RoboDK station: Bench V1 cell v4.rdk

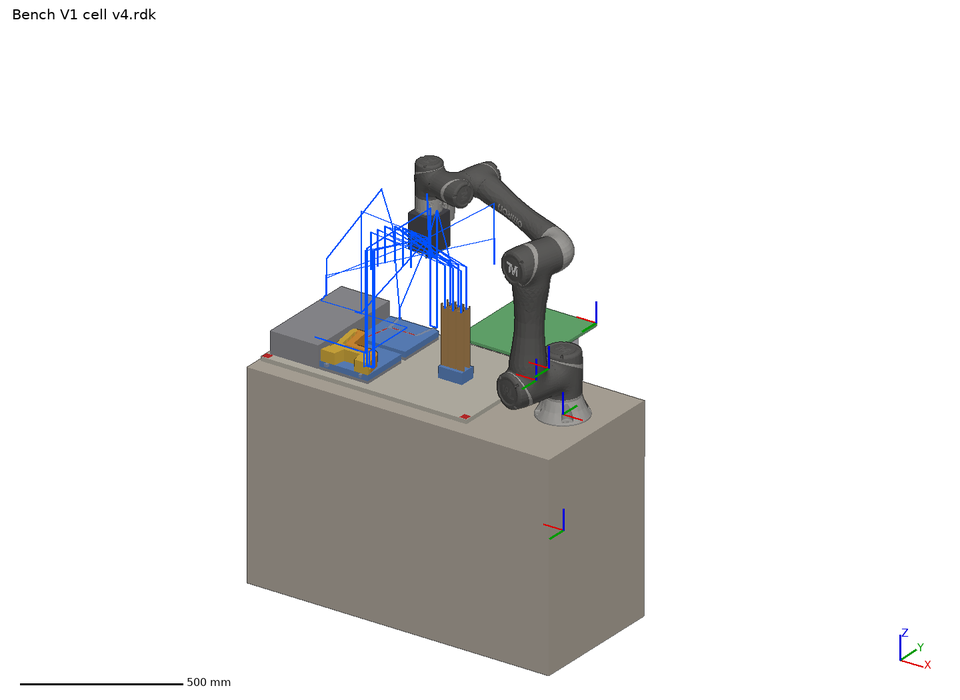
[picture v0: the station drawn from its stored meshes, robots at their saved joint values, targets as dots, program paths as lines]
Station Bench V1 cell v4 (saved by RoboDK 6.1.1). Poses are relative to the parent item; angles as X-Y-Z fixed-axis rotations.
Station parameters (name, value as stored): IO_0, 0
  - frame Cell at (0, 0, 0) mm
    - frame Work plate at (-206.44, 152.99, -4.46) mm, rotated rx -0.03 ry -0.07 rz -179.98 deg
      - frame Ground base at (0, -67, 15) mm
        - object Table at (0, 0, 0) mm, size 1130 x 510 x 735 mm
        - object Ground base plate at (0, 0, 0) mm, size 770 x 440 x 15 mm, geometry from ground_base_split.stl
        - object Vision square 1 at (3, 3, 0) mm, size 25 x 25 x 0.5 mm, geometry from vision_square.stl
        - object Vision square 2 at (742, 3, 0) mm, size 25 x 25 x 0.5 mm, geometry from vision_square.stl
        - object Vision square 3 at (3, 412, 0) mm, size 25 x 25 x 0.5 mm, geometry from vision_square.stl
        - object Vision square 4 at (742, 412, 0) mm, size 25 x 25 x 0.5 mm, geometry from vision_square.stl
        - object Base A riser at (480, 120, 10) mm, size 180 x 180 x 10 mm
        - object Base A at (480, 120, 10) mm, size 180 x 180 x 20 mm, geometry from base_a.stl
        - object Base B riser at (480, 320, 10) mm, size 180 x 180 x 10 mm
        - object Base B at (480, 320, 10) mm, size 180 x 180 x 20 mm, geometry from base_b.stl
        - object Plank jig at (150, 190, 0) mm, size 90 x 60 x 40 mm, geometry from plank_jig.stl
        - object Parking pad at (665, 220, 80) mm, size 180 x 380 x 80 mm, geometry from parking_pad.stl
        - frame AMR at (60, -340, 0) mm
          - object AMR plate at (0, 0, 0) mm, size 300 x 320 x 10 mm
          - object AMR top module at (0, 0, 0) mm, size 220 x 240 x 372 mm
          - frame Omron LD-250 Base at (150, -40, -765) mm
            - robot AMR LD-250: 4 axes
                joint limits [-10000, -10000, -10, -3600] to [10000, 10000, 10, 3600]; home [0, 0, 0, 0]; saved at [0, 0, 0, 0]
        - target Home (Cartesian target) at (295, 220, 380) mm, rotated rx 180 ry 0 rz 0 deg; joints [-14.089, 2.917, -80.099, -12.747, -90.01, 75.887] of Omron TM5-900
        - target guide B-A pick out low (Cartesian target) at (383, 390, 50) mm, rotated rx 0 ry 90 rz 0 deg; joints [8.389, -22.724, -132.74, -24.469, 98.365, 89.963] of Omron TM5-900
        - target guide B-A pick out (Cartesian target) at (383, 390, 450) mm, rotated rx 0 ry 90 rz 0 deg; joints [8.433, 10.061, -100.143, -89.851, 98.409, 89.963] of Omron TM5-900
        - target guide B-A via (Cartesian target) at (295, 220, 450) mm, rotated rx 0 ry 90 rz 0 deg; joints [-32.59, 30.389, -113.158, -97.152, 57.386, 90.016] of Omron TM5-900
        - target guide B-A centre (Cartesian target) at (295, 220, 450) mm, rotated rx 180 ry 0 rz 0 deg; joints [-14.088, -0.071, -66.923, -22.935, -90.01, 75.888] of Omron TM5-900
        - target guide B-A wrist ready (Cartesian target) at (295, 220, 450) mm, rotated rx -104.58 ry -32.51 rz -35.37 deg; joints [-50.735, 20.512, -106.829, -34.479, -14.275, 24.972] of Omron TM5-900
        - target guide B-A wrist swapped (joint target) at (338.92, 166.34, 566.06) mm, rotated rx -75.5 ry -32.53 rz -66.11 deg; joints [-50.735, 20.512, -106.829, -34.479, 14.275, 24.972] of Omron TM5-900
        - target guide B-A via (Cartesian target) at (295, 220, 450) mm, rotated rx 0 ry 90 rz 0 deg; joints [-32.59, 30.389, -113.158, -97.152, 57.386, 90.016] of Omron TM5-900
        - target guide B-A pick (Cartesian target) at (408, 390, 50) mm, rotated rx 0 ry 90 rz 0 deg; joints [7.812, -24.505, -129.214, -26.214, 97.788, 89.964] of Omron TM5-900
        - target guide B-A lift (Cartesian target) at (408, 390, 70) mm, rotated rx 0 ry 90 rz 0 deg; joints [7.814, -21.463, -128.95, -29.52, 97.79, 89.964] of Omron TM5-900
        - target guide B-A up (Cartesian target) at (408, 390, 450) mm, rotated rx 0 ry 90 rz 0 deg; joints [7.851, 6.883, -97.45, -89.366, 97.827, 89.964] of Omron TM5-900
        - target guide B-A across (Cartesian target) at (408, 50, 450) mm, rotated rx 0 ry 90 rz 0 deg; joints [-45.328, 6.909, -97.45, -89.364, 44.648, 90.04] of Omron TM5-900
        - target guide B-A place (Cartesian target) at (408, 50, 50) mm, rotated rx 0 ry -90 rz -180 deg; joints [-45.297, -24.479, -129.215, -26.212, 44.679, -89.96] of Omron TM5-900
        - target guide B-A over place (Cartesian target) at (408, 50, 450) mm, rotated rx 0 ry -90 rz -180 deg; joints [-45.328, 6.909, -97.45, -89.364, 44.648, -89.96] of Omron TM5-900
        - target guide B-A place approach (Cartesian target) at (408, 50, 90) mm, rotated rx 0 ry -90 rz -180 deg; joints [-45.3, -18.508, -128.521, -32.876, 44.676, -89.96] of Omron TM5-900
        - target guide B-A place out (Cartesian target) at (383, 50, 50) mm, rotated rx 0 ry -90 rz -180 deg; joints [-48.296, -22.696, -132.741, -24.463, 41.68, -89.952] of Omron TM5-900
        - target guide B-A place out up (Cartesian target) at (383, 50, 450) mm, rotated rx 0 ry -90 rz -180 deg; joints [-48.333, 10.089, -100.144, -89.845, 41.642, -89.952] of Omron TM5-900
        - target plank3 pick travel (Cartesian target) at (225, 205, 380) mm, rotated rx 180 ry 0 rz -90 deg; joints [-18.429, 12.369, -88.214, -14.084, -90.005, -198.454] of Omron TM5-900
        - target plank3 pick approach (Cartesian target) at (225, 205, 275) mm, rotated rx 180 ry 0 rz -90 deg; joints [-18.431, 14.063, -104.285, 0.293, -90.005, -198.455] of Omron TM5-900
        - target plank3 pick (Cartesian target) at (225, 205, 235) mm, rotated rx 180 ry 0 rz -90 deg; joints [-18.431, 13.759, -109.643, 5.956, -90.005, -198.455] of Omron TM5-900
        - target plank3 pick out (Cartesian target) at (225, 205, 295) mm, rotated rx 180 ry 0 rz -90 deg; joints [-18.43, 14.01, -101.456, -2.482, -90.005, -198.454] of Omron TM5-900
        - target plank3 pick up (Cartesian target) at (225, 205, 380) mm, rotated rx 180 ry 0 rz -90 deg; joints [-18.429, 12.369, -88.214, -14.084, -90.005, -198.454] of Omron TM5-900
        - target plank3 place travel (Cartesian target) at (507.27, 95.62, 380) mm, rotated rx 180 ry 0 rz -90 deg; joints [-19.585, -31.821, -35.961, -22.146, -90.003, -199.609] of Omron TM5-900
        - target plank3 above guide (Cartesian target) at (507.27, 95.62, 329.5) mm, rotated rx 180 ry 0 rz -90 deg; joints [-19.585, -28.774, -48.091, -13.064, -90.003, -199.609] of Omron TM5-900
        - target plank3 place (Cartesian target) at (507.27, 95.62, 254.5) mm, rotated rx 180 ry 0 rz -90 deg; joints [-19.585, -27.192, -61.018, -1.719, -90.003, -199.609] of Omron TM5-900
        - target plank3 push approach (Cartesian target) at (507.27, 95.62, 289.5) mm, rotated rx 180 ry 0 rz -90 deg; joints [-19.585, -27.6, -55.517, -6.811, -90.003, -199.609] of Omron TM5-900
        - target plank3 push (Cartesian target) at (507.27, 95.62, 269.5) mm, rotated rx 180 ry 0 rz -90 deg; joints [-19.585, -27.304, -58.757, -3.867, -90.003, -199.609] of Omron TM5-900
        - target plank3 push out (Cartesian target) at (507.27, 95.62, 289.5) mm, rotated rx 180 ry 0 rz -90 deg; joints [-19.585, -27.6, -55.517, -6.811, -90.003, -199.609] of Omron TM5-900
        - target plank3 place up (Cartesian target) at (507.27, 95.62, 380) mm, rotated rx 180 ry 0 rz -90 deg; joints [-19.585, -31.821, -35.961, -22.146, -90.003, -199.609] of Omron TM5-900
        - target plank6 pick travel (Cartesian target) at (225, 235, 380) mm, rotated rx 180 ry 0 rz -90 deg; joints [-14.439, 12.367, -88.214, -14.082, -90.01, -194.463] of Omron TM5-900
        - target plank6 pick approach (Cartesian target) at (225, 235, 275) mm, rotated rx 180 ry 0 rz -90 deg; joints [-14.441, 14.061, -104.285, 0.295, -90.01, -194.465] of Omron TM5-900
        - target plank6 pick (Cartesian target) at (225, 235, 235) mm, rotated rx 180 ry 0 rz -90 deg; joints [-14.442, 13.757, -109.644, 5.958, -90.01, -194.466] of Omron TM5-900
        - target plank6 pick out (Cartesian target) at (225, 235, 295) mm, rotated rx 180 ry 0 rz -90 deg; joints [-14.441, 14.009, -101.457, -2.481, -90.01, -194.465] of Omron TM5-900
        - target plank6 pick up (Cartesian target) at (225, 235, 380) mm, rotated rx 180 ry 0 rz -90 deg; joints [-14.439, 12.367, -88.214, -14.082, -90.01, -194.463] of Omron TM5-900
        - target plank6 place travel (Cartesian target) at (542.12, 175.18, 380) mm, rotated rx 180 ry 0 rz -10 deg; joints [-12.785, -37.947, -25.826, -26.156, -90.012, 87.191] of Omron TM5-900
        - target plank6 above guide (Cartesian target) at (542.12, 175.18, 329.5) mm, rotated rx 180 ry 0 rz -10 deg; joints [-12.785, -33.547, -40.655, -15.727, -90.012, 87.191] of Omron TM5-900
        - target plank6 place (Cartesian target) at (542.12, 175.18, 254.5) mm, rotated rx 180 ry 0 rz -10 deg; joints [-12.787, -31.253, -54.883, -3.793, -90.012, 87.189] of Omron TM5-900
        - target plank6 push approach (Cartesian target) at (542.12, 175.18, 289.5) mm, rotated rx 180 ry 0 rz -10 deg; joints [-12.786, -31.919, -48.939, -9.071, -90.012, 87.19] of Omron TM5-900
        - target plank6 push (Cartesian target) at (542.12, 175.18, 269.5) mm, rotated rx 180 ry 0 rz -10 deg; joints [-12.786, -31.466, -52.456, -6.008, -90.012, 87.19] of Omron TM5-900
        - target plank6 push out (Cartesian target) at (542.12, 175.18, 289.5) mm, rotated rx 180 ry 0 rz -10 deg; joints [-12.786, -31.919, -48.939, -9.071, -90.012, 87.19] of Omron TM5-900
        - target plank6 place up (Cartesian target) at (542.12, 175.18, 380) mm, rotated rx 180 ry 0 rz -10 deg; joints [-12.785, -37.947, -25.826, -26.156, -90.012, 87.191] of Omron TM5-900
        - target plank2 pick travel (Cartesian target) at (195, 205, 380) mm, rotated rx 180 ry 0 rz -90 deg; joints [-19.849, 16.424, -91.186, -15.166, -90.003, 160.127] of Omron TM5-900
        - target plank2 pick approach (Cartesian target) at (195, 205, 275) mm, rotated rx 180 ry 0 rz -90 deg; joints [-19.85, 18.419, -107.374, -0.973, -90.003, 160.126] of Omron TM5-900
        - target plank2 pick (Cartesian target) at (195, 205, 235) mm, rotated rx 180 ry 0 rz -90 deg; joints [-19.85, 18.235, -112.832, 4.668, -90.003, 160.126] of Omron TM5-900
        - target plank2 pick out (Cartesian target) at (195, 205, 295) mm, rotated rx 180 ry 0 rz -90 deg; joints [-19.85, 18.305, -104.507, -3.726, -90.003, 160.126] of Omron TM5-900
        - target plank2 pick up (Cartesian target) at (195, 205, 380) mm, rotated rx 180 ry 0 rz -90 deg; joints [-19.849, 16.424, -91.186, -15.166, -90.003, 160.127] of Omron TM5-900
        - target plank2 place travel (Cartesian target) at (447.3, 95.62, 380) mm, rotated rx 180 ry 0 rz -90 deg; joints [-21.345, -20.954, -52.182, -16.792, -90.001, 158.631] of Omron TM5-900
        - target plank2 above guide (Cartesian target) at (447.3, 95.62, 329.5) mm, rotated rx 180 ry 0 rz -90 deg; joints [-21.345, -19.166, -61.856, -8.907, -90.001, 158.631] of Omron TM5-900
        - target plank2 place (Cartesian target) at (447.3, 95.62, 254.5) mm, rotated rx 180 ry 0 rz -90 deg; joints [-21.345, -18.495, -73.245, 1.812, -90.001, 158.631] of Omron TM5-900
        - target plank2 push approach (Cartesian target) at (447.3, 95.62, 289.5) mm, rotated rx 180 ry 0 rz -90 deg; joints [-21.345, -18.55, -68.29, -3.088, -90.001, 158.631] of Omron TM5-900
        - target plank2 push (Cartesian target) at (447.3, 95.62, 269.5) mm, rotated rx 180 ry 0 rz -90 deg; joints [-21.345, -18.467, -71.191, -0.27, -90.001, 158.631] of Omron TM5-900
        - target plank2 push out (Cartesian target) at (447.3, 95.62, 289.5) mm, rotated rx 180 ry 0 rz -90 deg; joints [-21.345, -18.55, -68.29, -3.088, -90.001, 158.631] of Omron TM5-900
        - target plank2 place up (Cartesian target) at (447.3, 95.62, 380) mm, rotated rx 180 ry 0 rz -90 deg; joints [-21.345, -20.954, -52.182, -16.792, -90.001, 158.631] of Omron TM5-900
        - target plank5 pick travel (Cartesian target) at (195, 235, 380) mm, rotated rx 180 ry 0 rz -90 deg; joints [-15.56, 16.422, -91.186, -15.164, -90.008, 164.416] of Omron TM5-900
        - target plank5 pick approach (Cartesian target) at (195, 235, 275) mm, rotated rx 180 ry 0 rz -90 deg; joints [-15.562, 18.416, -107.374, -0.971, -90.008, 164.414] of Omron TM5-900
        - target plank5 pick (Cartesian target) at (195, 235, 235) mm, rotated rx 180 ry 0 rz -90 deg; joints [-15.563, 18.233, -112.832, 4.67, -90.008, 164.413] of Omron TM5-900
        - target plank5 pick out (Cartesian target) at (195, 235, 295) mm, rotated rx 180 ry 0 rz -90 deg; joints [-15.561, 18.303, -104.507, -3.724, -90.008, 164.415] of Omron TM5-900
        - target plank5 pick up (Cartesian target) at (195, 235, 380) mm, rotated rx 180 ry 0 rz -90 deg; joints [-15.56, 16.422, -91.186, -15.164, -90.008, 164.416] of Omron TM5-900
        - target plank5 place travel (Cartesian target) at (536.91, 145.66, 380) mm, rotated rx 180 ry 0 rz -10 deg; joints [-15.108, -37.171, -27.15, -25.608, -90.009, 84.868] of Omron TM5-900
        - target plank5 above guide (Cartesian target) at (536.91, 145.66, 329.5) mm, rotated rx 180 ry 0 rz -10 deg; joints [-15.109, -32.984, -41.552, -15.393, -90.009, 84.867] of Omron TM5-900
        - target plank5 place (Cartesian target) at (536.91, 145.66, 254.5) mm, rotated rx 180 ry 0 rz -10 deg; joints [-15.11, -30.786, -55.602, -3.541, -90.009, 84.866] of Omron TM5-900
        - target plank5 push approach (Cartesian target) at (536.91, 145.66, 289.5) mm, rotated rx 180 ry 0 rz -10 deg; joints [-15.109, -31.418, -49.717, -8.794, -90.009, 84.866] of Omron TM5-900
        - target plank5 push (Cartesian target) at (536.91, 145.66, 269.5) mm, rotated rx 180 ry 0 rz -10 deg; joints [-15.11, -30.985, -53.197, -5.747, -90.009, 84.866] of Omron TM5-900
        - target plank5 push out (Cartesian target) at (536.91, 145.66, 289.5) mm, rotated rx 180 ry 0 rz -10 deg; joints [-15.109, -31.418, -49.717, -8.794, -90.009, 84.866] of Omron TM5-900
        - target plank5 place up (Cartesian target) at (536.91, 145.66, 380) mm, rotated rx 180 ry 0 rz -10 deg; joints [-15.108, -37.171, -27.15, -25.608, -90.009, 84.868] of Omron TM5-900
        - target plank1 pick travel (Cartesian target) at (165, 205, 380) mm, rotated rx 180 ry 0 rz -90 deg; joints [-21.51, 20.489, -93.86, -16.558, -90.001, 158.466] of Omron TM5-900
        - target plank1 pick approach (Cartesian target) at (165, 205, 275) mm, rotated rx 180 ry 0 rz -90 deg; joints [-21.51, 22.877, -110.195, -2.609, -90.001, 158.466] of Omron TM5-900
        - target plank1 pick (Cartesian target) at (165, 205, 235) mm, rotated rx 180 ry 0 rz -90 deg; joints [-21.51, 22.858, -115.763, 2.976, -90.001, 158.466] of Omron TM5-900
        - target plank1 pick out (Cartesian target) at (165, 205, 295) mm, rotated rx 180 ry 0 rz -90 deg; joints [-21.51, 22.681, -107.284, -5.326, -90.001, 158.466] of Omron TM5-900
        - target plank1 pick up (Cartesian target) at (165, 205, 380) mm, rotated rx 180 ry 0 rz -90 deg; joints [-21.51, 20.489, -93.86, -16.558, -90.001, 158.466] of Omron TM5-900
        - target plank1 place travel (Cartesian target) at (477.29, 95.62, 380) mm, rotated rx 180 ry 0 rz -90 deg; joints [-20.428, -26.039, -44.868, -19.022, -90.002, 159.548] of Omron TM5-900
        - target plank1 above guide (Cartesian target) at (477.29, 95.62, 329.5) mm, rotated rx 180 ry 0 rz -90 deg; joints [-20.428, -23.785, -55.44, -10.703, -90.002, 159.548] of Omron TM5-900
        - target plank1 place (Cartesian target) at (477.29, 95.62, 254.5) mm, rotated rx 180 ry 0 rz -90 deg; joints [-20.428, -22.746, -67.427, 0.244, -90.002, 159.548] of Omron TM5-900
        - target plank1 push approach (Cartesian target) at (477.29, 95.62, 289.5) mm, rotated rx 180 ry 0 rz -90 deg; joints [-20.428, -22.948, -62.259, -4.722, -90.002, 159.548] of Omron TM5-900
        - target plank1 push (Cartesian target) at (477.29, 95.62, 269.5) mm, rotated rx 180 ry 0 rz -90 deg; joints [-20.428, -22.777, -65.292, -1.859, -90.002, 159.548] of Omron TM5-900
        - target plank1 push out (Cartesian target) at (477.29, 95.62, 289.5) mm, rotated rx 180 ry 0 rz -90 deg; joints [-20.428, -22.948, -62.259, -4.722, -90.002, 159.548] of Omron TM5-900
        - target plank1 place up (Cartesian target) at (477.29, 95.62, 380) mm, rotated rx 180 ry 0 rz -90 deg; joints [-20.428, -26.039, -44.868, -19.022, -90.002, 159.548] of Omron TM5-900
        - target plank4 pick travel (Cartesian target) at (165, 235, 380) mm, rotated rx 180 ry 0 rz -90 deg; joints [-16.873, 20.487, -93.86, -16.555, -90.006, 163.103] of Omron TM5-900
        - target plank4 pick approach (Cartesian target) at (165, 235, 275) mm, rotated rx 180 ry 0 rz -90 deg; joints [-16.875, 22.874, -110.196, -2.607, -90.006, 163.101] of Omron TM5-900
        - target plank4 pick (Cartesian target) at (165, 235, 235) mm, rotated rx 180 ry 0 rz -90 deg; joints [-16.876, 22.856, -115.763, 2.979, -90.006, 163.1] of Omron TM5-900
        - target plank4 pick out (Cartesian target) at (165, 235, 295) mm, rotated rx 180 ry 0 rz -90 deg; joints [-16.875, 22.679, -107.285, -5.323, -90.006, 163.101] of Omron TM5-900
        - target plank4 pick up (Cartesian target) at (165, 235, 380) mm, rotated rx 180 ry 0 rz -90 deg; joints [-16.873, 20.487, -93.86, -16.555, -90.006, 163.103] of Omron TM5-900
        - target plank4 place travel (Cartesian target) at (531.7, 116.13, 380) mm, rotated rx 180 ry 0 rz -10 deg; joints [-17.431, -36.736, -27.886, -25.307, -90.006, 82.545] of Omron TM5-900
        - target plank4 above guide (Cartesian target) at (531.7, 116.13, 329.5) mm, rotated rx 180 ry 0 rz -10 deg; joints [-17.431, -32.661, -42.063, -15.205, -90.006, 82.545] of Omron TM5-900
        - target plank4 place (Cartesian target) at (531.7, 116.13, 254.5) mm, rotated rx 180 ry 0 rz -10 deg; joints [-17.432, -30.517, -56.013, -3.399, -90.006, 82.544] of Omron TM5-900
        - target plank4 push approach (Cartesian target) at (531.7, 116.13, 289.5) mm, rotated rx 180 ry 0 rz -10 deg; joints [-17.432, -31.13, -50.162, -8.637, -90.006, 82.544] of Omron TM5-900
        - target plank4 push (Cartesian target) at (531.7, 116.13, 269.5) mm, rotated rx 180 ry 0 rz -10 deg; joints [-17.432, -30.709, -53.62, -5.599, -90.006, 82.544] of Omron TM5-900
        - target plank4 push out (Cartesian target) at (531.7, 116.13, 289.5) mm, rotated rx 180 ry 0 rz -10 deg; joints [-17.432, -31.13, -50.162, -8.637, -90.006, 82.544] of Omron TM5-900
        - target plank4 place up (Cartesian target) at (531.7, 116.13, 380) mm, rotated rx 180 ry 0 rz -10 deg; joints [-17.431, -36.736, -27.886, -25.307, -90.006, 82.545] of Omron TM5-900
        - target guide A-B pick out low (Cartesian target) at (383, 50, 50) mm, rotated rx 0 ry -90 rz -180 deg; joints [-48.296, -22.696, -132.741, -24.463, 41.68, -89.952] of Omron TM5-900
        - target guide A-B pick out (Cartesian target) at (383, 50, 450) mm, rotated rx 0 ry -90 rz -180 deg; joints [-48.333, 10.089, -100.144, -89.845, 41.642, -89.952] of Omron TM5-900
        - target guide A-B via (Cartesian target) at (295, 220, 450) mm, rotated rx 0 ry -90 rz -180 deg; joints [-32.59, 30.389, -113.158, -97.152, 57.386, -89.984] of Omron TM5-900
        - target guide A-B centre (Cartesian target) at (295, 220, 450) mm, rotated rx 180 ry 0 rz -10 deg; joints [-14.088, -0.071, -66.923, -22.935, -90.01, 85.888] of Omron TM5-900
        - target guide A-B wrist ready (Cartesian target) at (295, 220, 450) mm, rotated rx -103.31 ry -22.81 rz -38.08 deg; joints [-50.735, 20.512, -106.829, -34.479, -14.275, 34.972] of Omron TM5-900
        - target guide A-B wrist swapped (joint target) at (338.92, 166.34, 566.06) mm, rotated rx -76.76 ry -22.82 rz -63.41 deg; joints [-50.735, 20.512, -106.829, -34.479, 14.275, 34.972] of Omron TM5-900
        - target guide A-B via (Cartesian target) at (295, 220, 450) mm, rotated rx 0 ry -90 rz -180 deg; joints [-32.59, 30.389, -113.158, -97.152, 57.386, -89.984] of Omron TM5-900
        - target guide A-B pick (Cartesian target) at (408, 50, 50) mm, rotated rx 0 ry -90 rz -180 deg; joints [-45.297, -24.479, -129.215, -26.212, 44.679, -89.96] of Omron TM5-900
        - target guide A-B lift (Cartesian target) at (408, 50, 70) mm, rotated rx 0 ry -90 rz -180 deg; joints [-45.298, -21.437, -128.951, -29.518, 44.678, -89.96] of Omron TM5-900
        - target guide A-B up (Cartesian target) at (408, 50, 450) mm, rotated rx 0 ry -90 rz -180 deg; joints [-45.328, 6.909, -97.45, -89.364, 44.648, -89.96] of Omron TM5-900
        - target guide A-B across (Cartesian target) at (408, 390, 450) mm, rotated rx 0 ry -90 rz -180 deg; joints [7.851, 6.883, -97.45, -89.366, 97.827, -90.036] of Omron TM5-900
        - target guide A-B place (Cartesian target) at (408, 390, 50) mm, rotated rx 0 ry 90 rz 0 deg; joints [7.812, -24.505, -129.214, -26.214, 97.788, 89.964] of Omron TM5-900
        - target guide A-B over place (Cartesian target) at (408, 390, 450) mm, rotated rx 0 ry 90 rz 0 deg; joints [7.851, 6.883, -97.45, -89.366, 97.827, 89.964] of Omron TM5-900
        - target guide A-B place approach (Cartesian target) at (408, 390, 90) mm, rotated rx 0 ry 90 rz 0 deg; joints [7.816, -18.534, -128.521, -32.878, 97.792, 89.964] of Omron TM5-900
        - target guide A-B place out (Cartesian target) at (383, 390, 50) mm, rotated rx 0 ry 90 rz 0 deg; joints [8.389, -22.724, -132.74, -24.469, 98.365, 89.963] of Omron TM5-900
        - target guide A-B place out up (Cartesian target) at (383, 390, 450) mm, rotated rx 0 ry 90 rz 0 deg; joints [8.433, 10.061, -100.143, -89.851, 98.409, 89.963] of Omron TM5-900
        - target sub pick (Cartesian target) at (540.8, 23.3, 22) mm, rotated rx -120 ry 0 rz 9.93 deg; joints [-36.46, -73.895, -17.579, -49.907, -53.325, 25.436] of Omron TM5-900
        - target sub pick approach (Cartesian target) at (540.8, 23.3, 62) mm, rotated rx -120 ry 0 rz 9.93 deg; joints [-36.46, -74.48, -10.825, -56.077, -53.326, 25.435] of Omron TM5-900
        - target sub via (Cartesian target) at (295, 220, 450) mm, rotated rx -120 ry 0 rz 9.93 deg; joints [-35.279, -15.9, -56.713, -68.206, -52.406, 26.366] of Omron TM5-900
        - target sub centre (Cartesian target) at (295, 220, 450) mm, rotated rx 0 ry 90 rz 0 deg; joints [-32.59, 30.389, -113.158, -97.152, 57.386, 90.016] of Omron TM5-900
        - target sub start wrist ready (Cartesian target) at (295, 220, 450) mm, rotated rx 0 ry 90 rz 25 deg; joints [-50.744, 22.08, -108.673, -93.281, 14.232, 90.072] of Omron TM5-900
        - target sub start wrist swapped (joint target) at (209.75, 324.41, 449.85) mm, rotated rx 0 ry 90 rz 53.46 deg; joints [-50.744, 22.08, -108.673, -93.281, -14.231, 90.072] of Omron TM5-900
        - target sub to middle (joint target) at (430, 220, 450) mm, rotated rx -120 ry 0 rz 9.93 deg; joints [-28.865, -39.901, -20.638, -76.748, -47.557, 31.854] of Omron TM5-900
        - target sub wrist ready (Cartesian target) at (430, 220, 450) mm, rotated rx -98.01 ry -11.5 rz -23.96 deg; joints [-37.562, -12.266, -74.557, -59.684, -14.31, 20.984] of Omron TM5-900
        - target sub wrist swapped (joint target) at (519.65, 151.03, 524.65) mm, rotated rx -82.03 ry -11.51 rz -51.2 deg; joints [-37.562, -12.266, -74.557, -59.684, 14.31, 20.983] of Omron TM5-900
        - target sub place (Cartesian target) at (540.8, 416.7, 267) mm, rotated rx 60 ry 0 rz -9.93 deg; joints [20.85, -81.114, -28.985, 61.645, 138.058, 40.091] of Omron TM5-900
        - target sub above guide (Cartesian target) at (540.8, 416.7, 342) mm, rotated rx 60 ry 0 rz -9.93 deg; joints [20.854, -74.914, -30.845, 57.309, 138.056, 40.086] of Omron TM5-900
        - target sub flipped (Cartesian target) at (540.8, 416.7, 387) mm, rotated rx 60 ry 0 rz -9.93 deg; joints [20.856, -72.042, -30.214, 53.807, 138.054, 40.083] of Omron TM5-900
        - target sub place out (Cartesian target) at (544.53, 438.03, 254.5) mm, rotated rx 60 ry 0 rz -9.93 deg; joints [22.031, -87.305, -18.07, 57.884, 137.268, 38.788] of Omron TM5-900
        - target sub clear (Cartesian target) at (394.53, 438.03, 254.5) mm, rotated rx 60 ry 0 rz -9.93 deg; joints [26.213, -65.651, -65.413, 86.666, 134.358, 34.476] of Omron TM5-900
        - target sub back to middle (Cartesian target) at (295, 220, 450) mm, rotated rx 60 ry 0 rz -9.93 deg; joints [11.416, -24.337, -106.582, 73.148, 143.748, 52.064] of Omron TM5-900
        - target inner pick out low (Cartesian target) at (383, 385, 50) mm, rotated rx 0 ry 90 rz 0 deg; joints [7.543, -22.535, -133.111, -24.287, 97.519, 89.964] of Omron TM5-900
        - target inner pick out (Cartesian target) at (383, 385, 450) mm, rotated rx 0 ry 90 rz 0 deg; joints [7.586, 10.4, -100.419, -89.914, 97.562, 89.964] of Omron TM5-900
        - target inner via (Cartesian target) at (295, 220, 450) mm, rotated rx 0 ry 90 rz 0 deg; joints [-32.59, 30.389, -113.158, -97.152, 57.386, 90.016] of Omron TM5-900
        - target inner pick (Cartesian target) at (408, 385, 50) mm, rotated rx 0 ry 90 rz 0 deg; joints [7.02, -24.326, -129.566, -26.041, 96.996, 89.965] of Omron TM5-900
        - target inner out 1 (Cartesian target) at (400.12, 383.61, 50) mm, rotated rx 0 ry 90 rz 0 deg; joints [6.951, -23.709, -130.79, -25.435, 96.927, 89.965] of Omron TM5-900
        - target inner out 2 (Cartesian target) at (400.12, 383.61, 100) mm, rotated rx 0 ry 90 rz 0 deg; joints [6.956, -16.102, -129.798, -34.033, 96.932, 89.965] of Omron TM5-900
        - target inner out 3 (Cartesian target) at (400.12, 185, 100) mm, rotated rx 0 ry 90 rz 0 deg; joints [-27.469, -12.242, -135.436, -32.248, 62.507, 90.008] of Omron TM5-900
        - target inner out 4 (Cartesian target) at (595.12, 185, 100) mm, rotated rx 0 ry 90 rz 0 deg; joints [-17.159, -31.708, -103.725, -44.497, 72.816, 89.994] of Omron TM5-900
        - target inner place out (Cartesian target) at (570.12, 185, 100) mm, rotated rx 0 ry 90 rz 0 deg; joints [-18.024, -29.251, -108.074, -42.606, 71.952, 89.995] of Omron TM5-900
        - target inner place out up (Cartesian target) at (570.12, 185, 450) mm, rotated rx 0 ry 90 rz 0 deg; joints [-18.021, -10.311, -79.681, -89.938, 71.955, 89.995] of Omron TM5-900
        - target outer pick out low (Cartesian target) at (383, 395, 50) mm, rotated rx 0 ry 90 rz 0 deg; joints [9.228, -22.917, -132.359, -24.656, 99.204, 89.962] of Omron TM5-900
        - target outer pick out (Cartesian target) at (383, 395, 450) mm, rotated rx 0 ry 90 rz 0 deg; joints [9.272, 9.714, -99.859, -89.788, 99.248, 89.962] of Omron TM5-900
        - target outer via (Cartesian target) at (295, 220, 450) mm, rotated rx 0 ry 90 rz 0 deg; joints [-32.59, 30.389, -113.158, -97.152, 57.386, 90.016] of Omron TM5-900
        - target outer pick (Cartesian target) at (408, 395, 50) mm, rotated rx 0 ry 90 rz 0 deg; joints [8.597, -24.687, -128.854, -26.392, 98.573, 89.963] of Omron TM5-900
        - target outer out 1 (Cartesian target) at (408, 403, 50) mm, rotated rx 0 ry 90 rz 0 deg; joints [9.838, -24.988, -128.259, -26.685, 99.814, 89.962] of Omron TM5-900
        - target outer out 2 (Cartesian target) at (408, 403, 100) mm, rotated rx 0 ry 90 rz 0 deg; joints [9.844, -17.727, -127.303, -34.903, 99.82, 89.962] of Omron TM5-900
        - target outer out 3 (Cartesian target) at (593, 403, 100) mm, rotated rx 0 ry 90 rz 0 deg; joints [6.531, -34.487, -98.753, -46.694, 96.507, 89.965] of Omron TM5-900
        - target outer place out (Cartesian target) at (403, 403, 100) mm, rotated rx 0 ry 90 rz 0 deg; joints [9.979, -17.281, -127.995, -34.656, 99.955, 89.961] of Omron TM5-900
        - target outer place out up (Cartesian target) at (403, 403, 450) mm, rotated rx 0 ry 90 rz 0 deg; joints [10.016, 6.655, -97.252, -89.336, 99.991, 89.961] of Omron TM5-900
        - target bench pick out low (Cartesian target) at (540.8, 416.7, 287) mm, rotated rx 180 ry 0 rz -9.93 deg; joints [5.685, -36.085, -42.671, -11.181, -90.033, 105.587] of Omron TM5-900
        - target bench pick out (Cartesian target) at (540.8, 416.7, 322) mm, rotated rx 180 ry 0 rz -9.93 deg; joints [5.687, -37.936, -34.58, -17.421, -90.033, 105.589] of Omron TM5-900
        - target bench via (Cartesian target) at (295, 220, 450) mm, rotated rx 180 ry 0 rz -9.93 deg; joints [-14.088, -0.071, -66.923, -22.935, -90.01, 85.814] of Omron TM5-900
        - target bench centre (Cartesian target) at (295, 220, 450) mm, rotated rx 0 ry 90 rz 0 deg; joints [-32.59, 30.389, -113.158, -97.152, 57.386, 90.016] of Omron TM5-900
        - target bench wrist ready (Cartesian target) at (295, 220, 450) mm, rotated rx 0 ry 90 rz 25 deg; joints [-50.744, 22.08, -108.673, -93.281, 14.232, 90.072] of Omron TM5-900
        - target bench wrist swapped (joint target) at (209.75, 324.41, 449.85) mm, rotated rx 0 ry 90 rz 53.46 deg; joints [-50.744, 22.08, -108.673, -93.281, -14.231, 90.072] of Omron TM5-900
        - target bench via (Cartesian target) at (295, 220, 450) mm, rotated rx 180 ry 0 rz -9.93 deg; joints [-14.088, -0.071, -66.923, -22.935, -90.01, 85.814] of Omron TM5-900
        - target bench pick (Cartesian target) at (540.8, 416.7, 262) mm, rotated rx 180 ry 0 rz -9.93 deg; joints [5.684, -35.332, -47.421, -7.184, -90.033, 105.586] of Omron TM5-900
        - target bench lift (Cartesian target) at (540.8, 416.7, 332) mm, rotated rx 180 ry 0 rz -9.93 deg; joints [5.687, -38.707, -31.813, -19.417, -90.033, 105.589] of Omron TM5-900
        - target bench over AMR (Cartesian target) at (265.8, -89.8, 332) mm, rotated rx 180 ry 0 rz -9.93 deg; joints [-45.79, -4.744, -79.08, -6.111, -89.971, 54.112] of Omron TM5-900
        - target bench down (Cartesian target) at (265.8, -89.8, 243) mm, rotated rx 180 ry 0 rz -9.93 deg; joints [-45.786, -4.767, -91.487, 6.319, -89.971, 54.116] of Omron TM5-900
        - target bench place out (Cartesian target) at (265.8, -89.8, 283) mm, rotated rx 180 ry 0 rz -9.93 deg; joints [-45.788, -4.436, -86.256, 0.758, -89.971, 54.114] of Omron TM5-900
        - target bench place out up (Cartesian target) at (265.8, -89.8, 450) mm, rotated rx 180 ry 0 rz -9.93 deg; joints [-45.797, -9.125, -57.026, -23.783, -89.971, 54.106] of Omron TM5-900
        - target back to middle (Cartesian target) at (295, 220, 450) mm, rotated rx -180 ry 0 rz -9.93 deg; joints [-14.088, -0.071, -66.923, -22.935, -90.01, 85.814] of Omron TM5-900
        - object Guide inner at (480, 320, 90) mm, rotated rx 180 ry 0 rz 0 deg, size 158.3 x 160 x 40 mm, geometry from guide_inner.stl
        - object Guide outer at (480, 320, 90) mm, rotated rx 180 ry 0 rz 0 deg, size 177.7 x 180 x 40 mm, geometry from guide_outer.stl
        - object frame1 at (477.29, 93.12, 144.5) mm, rotated rx 0 ry 0 rz -90 deg, size 174.7 x 141.9 x 10 mm, geometry from frame.stl
        - object frame2 at (477.29, 346.88, -95.5) mm, rotated rx 180 ry 0 rz 90 deg, size 174.7 x 141.9 x 10 mm, geometry from frame.stl
        - object plank1 at (165, 207.5, 125) mm, rotated rx 90 ry 0 rz 0 deg, size 25 x 250 x 5 mm, geometry from plank_body.stl
        - object plank2 at (195, 207.5, 125) mm, rotated rx 90 ry 0 rz 0 deg, size 25 x 250 x 5 mm, geometry from plank_body.stl
        - object plank3 at (225, 207.5, 125) mm, rotated rx 90 ry 0 rz 0 deg, size 25 x 250 x 5 mm, geometry from plank_body.stl
        - object plank4 at (165, 237.5, 125) mm, rotated rx 90 ry 0 rz 0 deg, size 25 x 250 x 5 mm, geometry from plank_body.stl
        - object plank5 at (195, 237.5, 125) mm, rotated rx 90 ry 0 rz 0 deg, size 25 x 250 x 5 mm, geometry from plank_body.stl
        - object plank6 at (225, 237.5, 125) mm, rotated rx 90 ry 0 rz 0 deg, size 25 x 250 x 5 mm, geometry from plank_body.stl
        - object piece A1 at (477.29, 98.12, 144.5) mm, rotated rx 90 ry 0 rz 0 deg, size 21.4 x 10 x 5 mm, geometry from interface_piece.stl
        - object piece A2 at (447.3, 98.12, 144.5) mm, rotated rx 90 ry 0 rz 0 deg, size 21.4 x 10 x 5 mm, geometry from interface_piece.stl
        - object piece A3 at (507.27, 98.12, 144.5) mm, rotated rx 90 ry 0 rz 0 deg, size 21.4 x 10 x 5 mm, geometry from interface_piece.stl
        - object piece A4 at (529.24, 116.56, 144.5) mm, rotated rx 90 ry 0 rz 80 deg, size 21.4 x 10 x 5 mm, geometry from interface_piece.stl
        - object piece A5 at (534.45, 146.09, 144.5) mm, rotated rx 90 ry 0 rz 80 deg, size 21.4 x 10 x 5 mm, geometry from interface_piece.stl
        - object piece A6 at (539.66, 175.62, 144.5) mm, rotated rx 90 ry 0 rz 80 deg, size 21.4 x 10 x 5 mm, geometry from interface_piece.stl
        - object piece B1 at (477.29, 341.88, 144.5) mm, rotated rx 90 ry 0 rz -180 deg, size 21.4 x 10 x 5 mm, geometry from interface_piece.stl
        - object piece B2 at (447.3, 341.88, 144.5) mm, rotated rx 90 ry 0 rz -180 deg, size 21.4 x 10 x 5 mm, geometry from interface_piece.stl
        - object piece B3 at (507.27, 341.88, 144.5) mm, rotated rx 90 ry 0 rz -180 deg, size 21.4 x 10 x 5 mm, geometry from interface_piece.stl
        - object piece B4 at (529.24, 323.44, 144.5) mm, rotated rx 90 ry 0 rz 100 deg, size 21.4 x 10 x 5 mm, geometry from interface_piece.stl
        - object piece B5 at (534.45, 293.91, 144.5) mm, rotated rx 90 ry 0 rz 100 deg, size 21.4 x 10 x 5 mm, geometry from interface_piece.stl
        - object piece B6 at (539.66, 264.38, 144.5) mm, rotated rx 90 ry 0 rz 100 deg, size 21.4 x 10 x 5 mm, geometry from interface_piece.stl
    - frame Omron TM5-900 Base at (0, 0, 0) mm
      - robot Omron TM5-900: 6 axes, payload 4 kg, reach 900 mm, repeatability 0.05 mm, weight 22.6 kg
          modified DH rows (alpha deg, a mm, theta deg, d mm): 0, 0, 0, 145.2; 90, 0, 90, 0; 0, 429, 0, 0; 0, 411, -90, 122.3; -90, 0, 0, 106.5; 90, 0, 180, 114.15
          joint limits [-270, -180, -155, -180, -180, -270] to [270, 180, 155, 180, 180, 270]; home [0, 0, 90, -90, 90, 0]; saved at [-14.089, 2.917, -80.099, -12.747, -90.01, 75.887]
        - tool EGP, TCP at (0, 0, 160) mm, size 94 x 90 x 160 mm
  - program AssembleBench (342 instructions, listed below)
  - Python program Deliver (AMR) (listed below)
  - Python program Assemble and deliver (listed below)
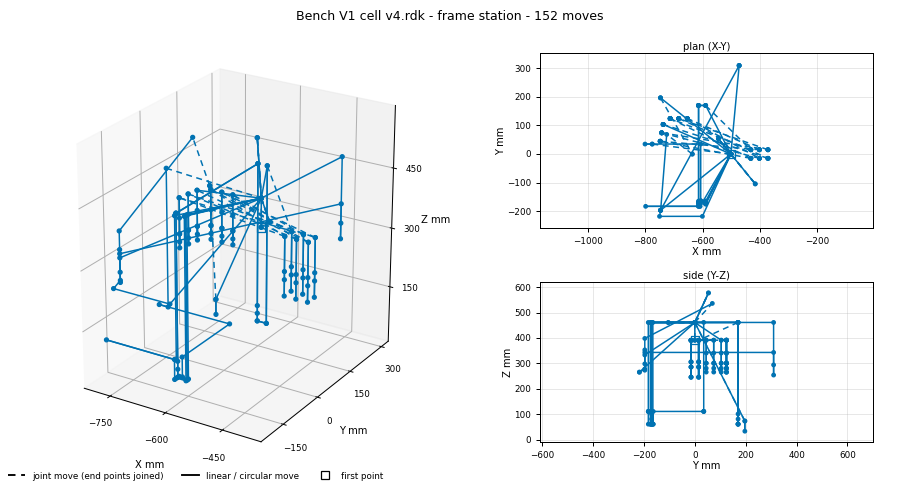
[picture p0: tool path of Bench V1 cell v4.rdk in frame station, 152 of 152 moves have a stored position in this frame; points joined in program order, loops and branches not executed]

--- program AssembleBench (robot Omron TM5-900) ---
  Simulation: parts to start
  Set Ref.: Ground base
  Set Tool: EGP
  Smooth(0)
  Set speed (100.0 mm/s)
  MoveJ (Home)
  MoveL (guide B-A centre)
  MoveL (guide B-A wrist ready)
  MoveJ (guide B-A wrist swapped)
  MoveL (guide B-A via)
  MoveL (guide B-A pick out)
  MoveL (guide B-A pick out low)
  Set speed (20.0 mm/s)
  Set IO_0=1
  Pause 300 ms
  MoveL (guide B-A pick)
  Set IO_0=0
  Pause 500 ms
  Simulation: attach Guide inner
  Simulation: attach Guide outer
  MoveL (guide B-A lift)
  Set speed (100.0 mm/s)
  MoveL (guide B-A up)
  MoveL (guide B-A across)
  MoveJ (guide B-A over place)
  MoveL (guide B-A place approach)
  Set speed (20.0 mm/s)
  MoveL (guide B-A place)
  Set IO_0=1
  Pause 500 ms
  Simulation: release guide B-A
  MoveL (guide B-A place out)
  Set speed (100.0 mm/s)
  MoveL (guide B-A place out up)
  MoveJ (plank3 pick travel)
  MoveL (plank3 pick approach)
  Set speed (20.0 mm/s)
  MoveL (plank3 pick)
  Set IO_0=1
  Pause 500 ms
  Simulation: attach plank3
  MoveL (plank3 pick out)
  Set speed (100.0 mm/s)
  MoveL (plank3 pick up)
  MoveJ (plank3 place travel)
  MoveL (plank3 above guide)
  Set speed (20.0 mm/s)
  MoveL (plank3 place)
  Set IO_0=0
  Pause 500 ms
  Simulation: release plank3
  MoveL (plank3 push approach)
  Set IO_0=1
  Pause 300 ms
  MoveL (plank3 push)
  MoveL (plank3 push out)
  Set IO_0=0
  Pause 300 ms
  Set speed (100.0 mm/s)
  MoveL (plank3 place up)
  MoveJ (plank6 pick travel)
  MoveL (plank6 pick approach)
  Set speed (20.0 mm/s)
  MoveL (plank6 pick)
  Set IO_0=1
  Pause 500 ms
  Simulation: attach plank6
  MoveL (plank6 pick out)
  Set speed (100.0 mm/s)
  MoveL (plank6 pick up)
  MoveJ (plank6 place travel)
  MoveL (plank6 above guide)
  Set speed (20.0 mm/s)
  MoveL (plank6 place)
  Set IO_0=0
  Pause 500 ms
  Simulation: release plank6
  MoveL (plank6 push approach)
  Set IO_0=1
  Pause 300 ms
  MoveL (plank6 push)
  MoveL (plank6 push out)
  Set IO_0=0
  Pause 300 ms
  Set speed (100.0 mm/s)
  MoveL (plank6 place up)
  MoveJ (plank2 pick travel)
  MoveL (plank2 pick approach)
  Set speed (20.0 mm/s)
  MoveL (plank2 pick)
  Set IO_0=1
  Pause 500 ms
  Simulation: attach plank2
  MoveL (plank2 pick out)
  Set speed (100.0 mm/s)
  MoveL (plank2 pick up)
  MoveJ (plank2 place travel)
  MoveL (plank2 above guide)
  Set speed (20.0 mm/s)
  MoveL (plank2 place)
  Set IO_0=0
  Pause 500 ms
  Simulation: release plank2
  MoveL (plank2 push approach)
  Set IO_0=1
  Pause 300 ms
  MoveL (plank2 push)
  MoveL (plank2 push out)
  Set IO_0=0
  Pause 300 ms
  Set speed (100.0 mm/s)
  MoveL (plank2 place up)
  MoveJ (plank5 pick travel)
  MoveL (plank5 pick approach)
  Set speed (20.0 mm/s)
  MoveL (plank5 pick)
  Set IO_0=1
  Pause 500 ms
  Simulation: attach plank5
  MoveL (plank5 pick out)
  Set speed (100.0 mm/s)
  MoveL (plank5 pick up)
  MoveJ (plank5 place travel)
  MoveL (plank5 above guide)
  Set speed (20.0 mm/s)
  MoveL (plank5 place)
  Set IO_0=0
  Pause 500 ms
  Simulation: release plank5
  MoveL (plank5 push approach)
  Set IO_0=1
  Pause 300 ms
  MoveL (plank5 push)
  MoveL (plank5 push out)
  Set IO_0=0
  Pause 300 ms
  Set speed (100.0 mm/s)
  MoveL (plank5 place up)
  MoveJ (plank1 pick travel)
  MoveL (plank1 pick approach)
  Set speed (20.0 mm/s)
  MoveL (plank1 pick)
  Set IO_0=1
  Pause 500 ms
  Simulation: attach plank1
  MoveL (plank1 pick out)
  Set speed (100.0 mm/s)
  MoveL (plank1 pick up)
  MoveJ (plank1 place travel)
  MoveL (plank1 above guide)
  Set speed (20.0 mm/s)
  MoveL (plank1 place)
  Set IO_0=0
  Pause 500 ms
  Simulation: release plank1
  MoveL (plank1 push approach)
  Set IO_0=1
  Pause 300 ms
  MoveL (plank1 push)
  MoveL (plank1 push out)
  Set IO_0=0
  Pause 300 ms
  Set speed (100.0 mm/s)
  MoveL (plank1 place up)
  MoveJ (plank4 pick travel)
  MoveL (plank4 pick approach)
  Set speed (20.0 mm/s)
  MoveL (plank4 pick)
  Set IO_0=1
  Pause 500 ms
  Simulation: attach plank4
  MoveL (plank4 pick out)
  Set speed (100.0 mm/s)
  MoveL (plank4 pick up)
  MoveJ (plank4 place travel)
  MoveL (plank4 above guide)
  Set speed (20.0 mm/s)
  MoveL (plank4 place)
  Set IO_0=0
  Pause 500 ms
  Simulation: release plank4
  MoveL (plank4 push approach)
  Set IO_0=1
  Pause 300 ms
  MoveL (plank4 push)
  MoveL (plank4 push out)
  Set IO_0=0
  Pause 300 ms
  Set speed (100.0 mm/s)
  MoveL (plank4 place up)
  MoveL (guide A-B centre)
  MoveL (guide A-B wrist ready)
  MoveJ (guide A-B wrist swapped)
  MoveL (guide A-B via)
  MoveL (guide A-B pick out)
  MoveL (guide A-B pick out low)
  Set speed (20.0 mm/s)
  Set IO_0=1
  Pause 300 ms
  MoveL (guide A-B pick)
  Set IO_0=0
  Pause 500 ms
  Simulation: attach Guide inner
  Simulation: attach Guide outer
  MoveL (guide A-B lift)
  Set speed (100.0 mm/s)
  MoveL (guide A-B up)
  MoveL (guide A-B across)
  MoveJ (guide A-B over place)
  MoveL (guide A-B place approach)
  Set speed (20.0 mm/s)
  MoveL (guide A-B place)
  Set IO_0=1
  Pause 500 ms
  Simulation: release guide A-B
  MoveL (guide A-B place out)
  Set speed (100.0 mm/s)
  MoveL (guide A-B place out up)
  MoveL (sub centre)
  MoveL (sub start wrist ready)
  MoveJ (sub start wrist swapped)
  MoveJ (sub via)
  MoveL (sub pick approach)
  Set speed (20.0 mm/s)
  MoveL (sub pick)
  Set IO_0=1
  Pause 500 ms
  Simulation: attach frame1
  Simulation: attach plank1
  Simulation: attach plank2
  Simulation: attach plank3
  Simulation: attach plank4
  Simulation: attach plank5
  Simulation: attach plank6
  Simulation: attach piece A1
  Simulation: attach piece A2
  Simulation: attach piece A3
  Simulation: attach piece A4
  Simulation: attach piece A5
  Simulation: attach piece A6
  MoveL (sub pick approach)
  Set speed (100.0 mm/s)
  MoveJ (sub to middle)
  MoveL (sub wrist ready)
  MoveJ (sub wrist swapped)
  MoveL (sub flipped)
  MoveL (sub above guide)
  Set speed (20.0 mm/s)
  MoveL (sub place)
  Set IO_0=0
  Pause 500 ms
  Simulation: release frame 1 with the planks
  MoveL (sub place out)
  MoveL (sub clear)
  MoveL (sub back to middle)
  Set speed (100.0 mm/s)
  MoveJ (inner via)
  MoveL (inner pick out)
  MoveL (inner pick out low)
  Set speed (20.0 mm/s)
  Set IO_0=1
  Pause 300 ms
  MoveL (inner pick)
  Set IO_0=0
  Pause 500 ms
  Simulation: attach Guide inner
  Set speed (20.0 mm/s)
  MoveL (inner out 1)
  MoveL (inner out 2)
  MoveL (inner out 3)
  MoveL (inner out 4)
  Set IO_0=1
  Pause 500 ms
  Simulation: release inner
  MoveL (inner place out)
  Set speed (100.0 mm/s)
  MoveL (inner place out up)
  MoveJ (outer via)
  MoveL (outer pick out)
  MoveL (outer pick out low)
  Set speed (20.0 mm/s)
  Set IO_0=1
  Pause 300 ms
  MoveL (outer pick)
  Set IO_0=0
  Pause 500 ms
  Simulation: attach Guide outer
  Set speed (20.0 mm/s)
  MoveL (outer out 1)
  MoveL (outer out 2)
  MoveL (outer out 3)
  Set IO_0=1
  Pause 500 ms
  Simulation: release outer
  MoveL (outer place out)
  Set speed (100.0 mm/s)
  MoveL (outer place out up)
  MoveL (bench centre)
  MoveL (bench wrist ready)
  MoveJ (bench wrist swapped)
  MoveL (bench via)
  MoveL (bench pick out)
  MoveL (bench pick out low)
  Set speed (20.0 mm/s)
  Set IO_0=0
  Pause 300 ms
  MoveL (bench pick)
  Set IO_0=1
  Pause 500 ms
  Simulation: attach frame1
  Simulation: attach frame2
  Simulation: attach plank1
  Simulation: attach plank2
  Simulation: attach plank3
  Simulation: attach plank4
  Simulation: attach plank5
  Simulation: attach plank6
  Simulation: attach piece A1
  Simulation: attach piece A2
  Simulation: attach piece A3
  Simulation: attach piece A4
  Simulation: attach piece A5
  Simulation: attach piece A6
  Simulation: attach piece B1
  Simulation: attach piece B2
  Simulation: attach piece B3
  Simulation: attach piece B4
  Simulation: attach piece B5
  Simulation: attach piece B6
  MoveL (bench lift)
  Set speed (100.0 mm/s)
  MoveL (bench over AMR)
  Set speed (20.0 mm/s)
  MoveL (bench down)
  Set IO_0=0
  Pause 500 ms
  Simulation: release bench
  MoveL (bench place out)
  Set speed (100.0 mm/s)
  MoveL (bench place out up)
  MoveL (back to middle)
  MoveJ (Home)

--- Python program Deliver (AMR) ---
"""The AMR drives the finished bench 2 m away along the table and comes back (RoboDK station script
"Deliver (AMR)").

    python robot_cell/amr_drive.py           also works from outside RoboDK

Needs only the robodk package. Everything under the station's "AMR" frame rides along: its plate,
top module and LD-250, and the bench once the robot program has set it down there (the program's
release puts the bench under the AMR frame).
"""
import time

from robodk import robolink, robomath

DISTANCE = 2000          # mm, along the ground base's x (away from the robot)
STEPS = 120              # per direction
PAUSE = 1.0              # s at the far end
OWN = ("AMR plate", "AMR top module")


def main():
    RDK = robolink.Robolink()
    amr = RDK.Item("AMR", robolink.ITEM_TYPE_FRAME)
    if not amr.Valid():
        raise SystemExit("no AMR in the open station")
    riding = [c for c in amr.Childs() if c.Type() == robolink.ITEM_TYPE_OBJECT and c.Name() not in OWN]
    home = amr.Pose()
    for out in (True, False):
        for i in range(1, STEPS + 1):
            s = i / STEPS if out else 1 - i / STEPS
            s = 0.5 - 0.5 * robomath.cos(robomath.pi * s)        # smooth start and stop
            amr.setPose(robomath.transl(DISTANCE * s, 0, 0) * home)
            RDK.Render(True)
            time.sleep(0.02)
        if out:
            time.sleep(PAUSE)
    amr.setPose(home)
    print(f"AMR drove {DISTANCE / 1000:.0f} m and back with {len(riding)} parts on its plate")


if __name__ == "__main__":
    main()

--- Python program Assemble and deliver ---
"""The whole cycle (station script "Assemble and deliver"): the robot program AssembleBench builds the
bench and sets it down on the AMR, then the AMR drives it 2 m along the table and back (amr_drive.py).

    python robot_cell/assemble_and_deliver.py      also works from outside RoboDK
"""
import time

from robodk import robolink

import amr_drive


def main():
    RDK = robolink.Robolink()
    prog = RDK.Item("AssembleBench", robolink.ITEM_TYPE_PROGRAM)
    if not prog.Valid():
        raise SystemExit("no AssembleBench in the open station")
    t0 = time.time()
    prog.RunProgram()
    time.sleep(1)
    while prog.Busy():
        time.sleep(0.2)
    print(f"AssembleBench done after {time.time() - t0:.0f} s (at the simulation speed)")
    amr_drive.main()


if __name__ == "__main__":
    main()
